// TwinCAT 3 PLC project ShowPLC
// ProgramVersion: 3.1.4026.27
// libraries:
//   Tc2_Standard, * (Beckhoff Automation GmbH)
//   Tc2_SUPS, * (Beckhoff Automation GmbH)
//   Tc2_System, * (Beckhoff Automation GmbH)
//   Tc2_Utilities, * (Beckhoff Automation GmbH)
//   Tc3_IotBase, * (Beckhoff Automation GmbH)
//   Tc3_IPCDiag, * (Beckhoff Automation GmbH)
//   Tc3_JsonXml, * (Beckhoff Automation GmbH)
// project tree:
//   DUTs/ E_JsonSection.TcDUT, E_LoadKind.TcDUT, ST_AcMeasurement.TcDUT, ST_BoxConfig.TcDUT, ST_FeedConfig.TcDUT, ST_GenericLoadConfig.TcDUT, ST_Harmonics.TcDUT, ST_LoadDemand.TcDUT, ST_MqttConfig.TcDUT
//   GVLs/ GVL_Config.TcGVL, GVL_Param.TcGVL, GVL_Persist.TcGVL
//   / PlcTask.TcTTO
//   POUs/ITFs/ I_FeedLoad.TcIO, I_JsonSource.TcIO, I_PowerMeter.TcIO
//   POUs/ MAIN.TcPOU
//   POUs/Power/ FB_EcPowerSupply.TcPOU, FB_GenericLoad.TcPOU, FB_PowerFeed.TcPOU, FB_PowerMeter_Sim.TcPOU, FB_SatelliteController.TcPOU
//   POUs/System/ FB_HostThermal.TcPOU (not stored), FB_ShowClock.TcPOU, FB_Telemetry.TcPOU, FB_IpcDiagnostics.TcPOU
//   POUs/Util/ F_CableFactor.TcPOU, F_CableLossW.TcPOU, F_CleanReal.TcPOU, F_CycleTimeS.TcPOU, F_FeedIdString.TcPOU, F_JsonHarmArray.TcPOU, F_JsonInt.TcPOU, F_JsonNum.TcPOU, F_JsonNumSigned.TcPOU, F_LowPass.TcPOU, F_PadNum.TcPOU, F_PowerAfterCable.TcPOU, F_WireOhms.TcPOU
// real-time tasks:
//   TASK PlcTask: cycle T#10ms, priority 20, ADS port 350
// I/O:
//   DEVICE Device 1 (EtherCAT), AmsNetId 192.168.30.11.2.1
//     Term 1 (EK1200) [EK1200-5000 EtherCAT Power supply (2A E-Bus)]
//       Term 10 (EL6070-0033) [EL6070-0033 1Ch. Licence key terminal, individual licences]
//       Term 2 (EL6090) [EL6090 Display terminal]
//       Term 3 (EL9227-5500) [EL9227-5500 Overcurrent protection 24V DC, 2Ch., max. 10A (sum), adjustable, extended functionalities]
//       Term 4 (EL9184) [EL9184 Potential Connection, 8 x 24V, 8 x Ground]
//       Term 5 (EL1259) [EL1259 8Ch. Dig Input 24V/8Ch. Dig. Output 24V with Multi-Time-Stamp]
//       Term 6 (EL3453-0100) [EL3453 3Ch. Power Measuring 100V]
//       Term 7 (EL3453-0100) [EL3453 3Ch. Power Measuring 100V]
//       Term 8 (EK1110) [EK1110 EtherCAT extension]
//     Box 17 (PS2001-2410) [PS2001-2410-1001 Power supply (24V, 10A, 1-phase)]
// variable links:
//   ShowPLC/ShowPLC Instance <-> Device 1 (EtherCAT)
//     PlcTask Inputs/MAIN.fbIpc.nEcCfgSlaves <-> InfoData/CfgSlaveCount
//     PlcTask Inputs/MAIN.fbIpc.nEcDevState <-> Inputs/DevState
//     PlcTask Inputs/MAIN.fbIpc.nEcSlaveCount <-> Inputs/SlaveCount

CONFIGURATION ShowPLC
    RESOURCE PLC ON TwinCAT3
        TASK PlcTask(INTERVAL := T#10ms, PRIORITY := 20);
        PROGRAM MAIN WITH PlcTask : MAIN;
    END_RESOURCE
END_CONFIGURATION

// ---- DUTs/E_JsonSection.TcDUT
{attribute 'qualified_only'}
{attribute 'strict'}
TYPE E_JsonSection :
(
    Circuit := 0,   // one row of the website's original circuits[] list
    Feed,           // one row of feeds[]
    Box,            // one row of boxes[]
    Load,           // one row of loads[]
    Diag,           // the body of the diag payload
    Harmonics       // one row of the harmonics payload
);
END_TYPE

// ---- DUTs/E_LoadKind.TcDUT
{attribute 'qualified_only'}
{attribute 'strict'}
TYPE E_LoadKind :
(
    Measured := 0,  // has its own measurement (box with an EtherCAT power supply)
    Rated,          // fixed rated power (generic load)
    Estimated       // gets a share of whatever is left on the feed (box without a supply)
);
END_TYPE

// ---- DUTs/ST_AcMeasurement.TcDUT
TYPE ST_AcMeasurement :
STRUCT
    bValid        : BOOL;   // the values below can be used
    bThdValid     : BOOL;   // the four THD values can be used
    fVoltsL1      : LREAL;  // V, L1 to ground
    fVoltsL2      : LREAL;  // V, L2 to ground
    fVoltsLL      : LREAL;  // V, L1 to L2
    fAmpsL1       : LREAL;  // A
    fAmpsL2       : LREAL;  // A
    fAmpsResidual : LREAL;  // A, summation transformer on the IN channel
    fPowerW       : LREAL;  // W,  P(L1) + P(L2)
    fApparentVA   : LREAL;  // VA, S(L1) + S(L2)
    fPowerFactor  : LREAL;  // 0..1
    fFrequencyHz  : LREAL;
    fThdVoltsL1   : LREAL;  // %
    fThdVoltsL2   : LREAL;  // %
    fThdAmpsL1    : LREAL;  // %
    fThdAmpsL2    : LREAL;  // %
END_STRUCT
END_TYPE

// ---- DUTs/ST_BoxConfig.TcDUT
TYPE ST_BoxConfig :
STRUCT
    sId               : STRING(20);     // slug of the name: lowercase letters, digits and '-'
    sControllerName   : STRING(40);     // exactly the label the website uses for this controller
    nFeedId           : INT := 1;       // index into GVL_Config.aFeeds
    bHasEcPowerSupply : BOOL;           // TRUE: live values come from the EtherCAT supply in the box
    nPixelCount       : UDINT;
    fMaxDcCurrent     : LREAL := 20.0;  // A
    fNominalDcVolts   : LREAL := 24.0;  // turns an estimated share into DC amps
    fPsuEfficiency    : LREAL := 0.95;  // DC power out / AC power in
    fWireLengthFt     : LREAL := 0.0;   // one-way length of the box's AC cable from where it branches off the feed
    nWireAwg          : INT := 12;      // AWG of one conductor, copper
END_STRUCT
END_TYPE

// ---- DUTs/ST_FeedConfig.TcDUT
TYPE ST_FeedConfig :
STRUCT
    sId           : STRING(20);     // short id used in the payloads: F1, F2
    sName         : STRING(40);
    fMaxAmps      : LREAL := 32.0;  // A per leg
    fWireLengthFt : LREAL := 0.0;   // one-way length of the infeed cable: meter to the point where the boxes branch off
    nWireAwg      : INT := 10;      // AWG of one conductor, copper
END_STRUCT
END_TYPE

// ---- DUTs/ST_GenericLoadConfig.TcDUT
TYPE ST_GenericLoadConfig :
STRUCT
    sId           : STRING(20);  // L1, L2, ...
    sName         : STRING(40);
    nFeedId       : INT := 1;    // index into GVL_Config.aFeeds
    fRatedPowerW  : LREAL;       // W at the load
    bEnabled      : BOOL;        // FALSE: counts as 0 W
    fWireLengthFt : LREAL := 0.0; // one-way length of the load's cable from where it branches off the feed
    nWireAwg      : INT := 14;   // AWG of one conductor, copper
END_STRUCT
END_TYPE

// ---- DUTs/ST_Harmonics.TcDUT
TYPE ST_Harmonics :
STRUCT
    bValid   : BOOL;
    aVoltsL1 : ARRAY[2..GVL_Param.HARMONIC_MAX_ORDER] OF LREAL;
    aVoltsL2 : ARRAY[2..GVL_Param.HARMONIC_MAX_ORDER] OF LREAL;
    aAmpsL1  : ARRAY[2..GVL_Param.HARMONIC_MAX_ORDER] OF LREAL;
    aAmpsL2  : ARRAY[2..GVL_Param.HARMONIC_MAX_ORDER] OF LREAL;
END_STRUCT
END_TYPE

// ---- DUTs/ST_LoadDemand.TcDUT
TYPE ST_LoadDemand :
STRUCT
    eKind        : E_LoadKind;  // how the feed treats this load
    fAcPowerW    : LREAL;       // W the load takes at the branch point, its own cable loss included. Measured and Rated loads only
    fCableLossW  : LREAL;       // W lost in the load's own cable. Measured and Rated: part of fAcPowerW. Estimated: from its current share
    fWeight      : LREAL;       // share weight: the pixel count. Estimated loads only
    fCableFactor : LREAL;       // 1/W: loss in the load's own cable = fCableFactor * (power at the load)^2. Estimated loads only
    bValid       : BOOL;        // FALSE: a measured load that is not reporting
END_STRUCT
END_TYPE

// ---- DUTs/ST_MqttConfig.TcDUT
TYPE ST_MqttConfig :
STRUCT
    bEnable     : BOOL := TRUE;
    sHost       : STRING(63) := '192.168.30.31';
    nPort       : UINT := 1883;
    sClientId   : STRING(63) := 'sfl-plc';
    sUser       : STRING(63) := 'plc';
    nKeepAliveS : UINT := 30;
    sTopicRoot  : STRING(63) := 'sfl/plc';
    tDashboard  : TIME := T#1S;
    tDiag       : TIME := T#5S;
    tHarmonics  : TIME := T#10S;
END_STRUCT
END_TYPE

// ---- GVLs/GVL_Config.TcGVL
{attribute 'qualified_only'}
VAR_GLOBAL
    // ---- development switches -------------------------------------------------
    bSimulateMeters   : BOOL := TRUE;   // TRUE: feeds read FB_PowerMeter_Sim. Set FALSE in step 4
    bSimulateSupplies : BOOL := TRUE;   // TRUE: supplies use their fSim values. Set FALSE in step 5

    // ---- model ----------------------------------------------------------------
    fFilterTimeS      : LREAL := 1.0;   // low-pass on feed and supply values before the split, seconds
    fVoltsPresentMin  : LREAL := 90.0;  // V per leg. Above this a feed counts as "on"

    // ---- cables ---------------------------------------------------------------
    // Every feed, box and load has a one-way cable length and an AWG. The loss in each cable is I^2 R
    // with that component's own current. Lengths below are placeholders until measured.
    fWireTempC          : LREAL := 20.0;   // conductor temperature for the resistance. Copper: +0.39 % per degree C
    fWireFactor         : LREAL := 1.0;    // 1.0 solid copper, about 1.03 stranded copper, about 1.6 aluminium
    fNominalAcVolts     : LREAL := 240.0;  // L1 to L2 at the loads. With the power factor it turns a load's power into the current in its cable
    fNominalPowerFactor : LREAL := 1.0;    // of the boxes and loads. Current = power / (volts * power factor)

    // ---- feeds ----------------------------------------------------------------
    aFeeds : ARRAY[1..GVL_Param.FEED_COUNT] OF ST_FeedConfig := [
        (sId := 'F1', sName := 'Feed 1', fMaxAmps := 32.0, fWireLengthFt := 100.0, nWireAwg := 10),
        (sId := 'F2', sName := 'Feed 2', fMaxAmps := 32.0, fWireLengthFt := 100.0, nWireAwg := 10)];

    // ---- satellite controller boxes ---------------------------------------------
    // sControllerName must match the website's label exactly. sId is its slug.
    // A box without an EtherCAT supply is estimated from its feed. Its DC amps use fNominalDcVolts (24 V unless set here).
    aBoxes : ARRAY[1..GVL_Param.BOX_COUNT] OF ST_BoxConfig := [
        (sId := 'porch',        sControllerName := 'Porch',        nFeedId := 1, bHasEcPowerSupply := FALSE, nPixelCount := 16325, fMaxDcCurrent := 80.0, fWireLengthFt := 50.0, nWireAwg := 12),
        (sId := 'metal-roof',   sControllerName := 'Metal Roof',   nFeedId := 2, bHasEcPowerSupply := FALSE, nPixelCount := 12820, fMaxDcCurrent := 80.0, fWireLengthFt := 50.0, nWireAwg := 12),
        (sId := 'center-gable', sControllerName := 'Center Gable', nFeedId := 1, bHasEcPowerSupply := TRUE,  nPixelCount := 2841,  fMaxDcCurrent := 20.0, fWireLengthFt := 50.0, nWireAwg := 12),
        (sId := 'courtyard',    sControllerName := 'Courtyard',    nFeedId := 1, bHasEcPowerSupply := TRUE,  nPixelCount := 452,   fMaxDcCurrent := 20.0, fWireLengthFt := 50.0, nWireAwg := 12),
        (sId := 'lawn-s-1',     sControllerName := 'Lawn S-1',     nFeedId := 1, bHasEcPowerSupply := TRUE,  nPixelCount := 1500,  fMaxDcCurrent := 20.0, fWireLengthFt := 50.0, nWireAwg := 12),
        (sId := 'lawn-s-2',     sControllerName := 'Lawn S-2',     nFeedId := 1, bHasEcPowerSupply := TRUE,  nPixelCount := 2541,  fMaxDcCurrent := 20.0, fWireLengthFt := 50.0, nWireAwg := 12),
        (sId := 'lawn-s-3',     sControllerName := 'Lawn S-3',     nFeedId := 2, bHasEcPowerSupply := TRUE,  nPixelCount := 6141,  fMaxDcCurrent := 20.0, fWireLengthFt := 50.0, nWireAwg := 12),
        (sId := 'lawn-n-1',     sControllerName := 'Lawn N-1',     nFeedId := 2, bHasEcPowerSupply := TRUE,  nPixelCount := 2450,  fMaxDcCurrent := 20.0, fWireLengthFt := 50.0, nWireAwg := 12),
        (sId := 'lawn-n-2',     sControllerName := 'Lawn N-2',     nFeedId := 2, bHasEcPowerSupply := TRUE,  nPixelCount := 4115,  fMaxDcCurrent := 20.0, fWireLengthFt := 50.0, nWireAwg := 12)];

    // ---- generic loads ------------------------------------------------------------
    // One row per GVL_Param.LOAD_COUNT.
    aLoads : ARRAY[1..GVL_Param.LOAD_COUNT] OF ST_GenericLoadConfig := [
        (sId := 'L1', sName := 'Metal Roof Floods', nFeedId := 2, fRatedPowerW := 20.0, bEnabled := TRUE, fWireLengthFt := 50.0, nWireAwg := 14),
        (sId := 'L2', sName := 'North Peak Floods', nFeedId := 2, fRatedPowerW := 20.0, bEnabled := TRUE, fWireLengthFt := 50.0, nWireAwg := 14),
        (sId := 'L3', sName := 'South Peak Floods', nFeedId := 2, fRatedPowerW := 20.0, bEnabled := TRUE, fWireLengthFt := 50.0, nWireAwg := 14)];

    // ---- EtherCAT power supplies (PS2001) -------------------------------------------
    // Info data scaling is not documented. 0.0 keeps the value out of the payload until it is checked in step 5.
    fPsuInfo1Scale : LREAL := 0.0;      // degrees C per count of "Info data 1" (temperature)
    fPsuInfo2Scale : LREAL := 0.0;      // volts per count of "Info data 2" (RMS input voltage)

    // ---- TF8330 -----------------------------------------------------------------------
    nTf8330FundamentalIndex : INT := 1; // element of aHarm1 that reads 100 (the fundamental): 1 if element 0 is the DC part, 0 if the arrays start at the fundamental, -1 if they start at the 2nd harmonic. Check in step 4

    // ---- MQTT ---------------------------------------------------------------------------
    stMqtt : ST_MqttConfig;             // defaults are in the type

    // ---- local time, for the midnight energy reset: US Central ---------------------------
    // UTC = local time + bias (minutes). wDay is the occurrence in the month: 1 = first, 2 = second, 5 = last.
    stTimeZone : ST_TimeZoneInformation := (
        bias         := 360,
        standardName := 'CST',
        standardDate := (wYear := 0, wMonth := 11, wDayOfWeek := 0, wDay := 1, wHour := 2),
        standardBias := 0,
        daylightName := 'CDT',
        daylightDate := (wYear := 0, wMonth := 3, wDayOfWeek := 0, wDay := 2, wHour := 2),
        daylightBias := -60);
END_VAR

// ---- GVLs/GVL_Param.TcGVL
{attribute 'qualified_only'}
VAR_GLOBAL CONSTANT
    FEED_COUNT         : INT := 2;
    BOX_COUNT          : INT := 9;
    LOAD_COUNT         : INT := 3;
    MAX_LOADS_PER_FEED : INT := GVL_Param.BOX_COUNT + GVL_Param.LOAD_COUNT;
    HARMONIC_MAX_ORDER : INT := 25;  // highest harmonic order kept and published. 2..63
END_VAR

// ---- GVLs/GVL_Persist.TcGVL
{attribute 'qualified_only'}
VAR_GLOBAL PERSISTENT
    sMqttPassword : STRING(63);                                  // empty = telemetry stays offline
    aEnergyWh     : ARRAY[1..GVL_Param.FEED_COUNT] OF LREAL;     // Wh per feed since local midnight
    nEnergyDay    : UDINT;                                       // local day number the counters belong to
END_VAR

// ---- POUs/ITFs/I_FeedLoad.TcIO
INTERFACE I_FeedLoad

// What this load asks of its feed this cycle.
METHOD GetDemand : ST_LoadDemand
END_METHOD

// The feed's answer to an Estimated load: its share of the unmeasured power.
METHOD SetShare
VAR_INPUT
    fShareW     : LREAL;  // W on the AC side
    bShareValid : BOOL;   // FALSE: the feed has no valid measurement
END_VAR
END_METHOD

END_INTERFACE

// ---- POUs/ITFs/I_JsonSource.TcIO
INTERFACE I_JsonSource

// Writes the keys of one JSON object. The caller opens and closes the object.
METHOD WriteJson
VAR_INPUT
    eSection : E_JsonSection;
END_VAR
VAR_IN_OUT
    fbJson : FB_JsonSaxWriter;
END_VAR
END_METHOD

END_INTERFACE

// ---- POUs/ITFs/I_PowerMeter.TcIO
INTERFACE I_PowerMeter

// Fills stMeas. Returns TRUE when the values are valid.
METHOD Read : BOOL
VAR_IN_OUT
    stMeas : ST_AcMeasurement;
END_VAR
END_METHOD

// Fills stHarm. Returns TRUE when the values are valid.
METHOD ReadHarmonics : BOOL
VAR_IN_OUT
    stHarm : ST_Harmonics;
END_VAR
END_METHOD

END_INTERFACE

// ---- POUs/MAIN.TcPOU
PROGRAM MAIN
VAR
    // Power model
    aFeeds     : ARRAY[1..GVL_Param.FEED_COUNT] OF FB_PowerFeed;
    aSimMeters : ARRAY[1..GVL_Param.FEED_COUNT] OF FB_PowerMeter_Sim;
    aBoxes     : ARRAY[1..GVL_Param.BOX_COUNT] OF FB_SatelliteController;
    aLoads     : ARRAY[1..GVL_Param.LOAD_COUNT] OF FB_GenericLoad;
    ipMeter    : I_PowerMeter;

    // Totals for the website's top-level keys
    fTotalPowerW   : LREAL;
    fTotalAmps     : LREAL;
    fEnergyTodayWh : LREAL;

    // Reporting
    fbClock     : FB_ShowClock;
    fbTelemetry : FB_Telemetry;
    fbIpc       : FB_IpcDiagnostics;

    // Persistent data
    bSavePersistent : BOOL;                    // set TRUE online to store GVL_Persist now
    fbSavePersist   : FB_WritePersistentData;

    i : INT;
    n : INT;
END_VAR

// Clock. On a new local day the energy counters start again
fbClock();
IF fbClock.bValid AND (fbClock.nLocalDay <> GVL_Persist.nEnergyDay) THEN
    FOR i := 1 TO GVL_Param.FEED_COUNT DO
        GVL_Persist.aEnergyWh[i] := 0.0;
    END_FOR
    GVL_Persist.nEnergyDay := fbClock.nLocalDay;
END_IF

// Feeds: read the meter, filter, cable loss, start a new load list
FOR i := 1 TO GVL_Param.FEED_COUNT DO
    ipMeter := aSimMeters[i];
    aFeeds[i](stCfg := GVL_Config.aFeeds[i], ipMeter := ipMeter, fEnergyWh := GVL_Persist.aEnergyWh[i]);
END_FOR

// Boxes and generic loads: update, then report to their feed
FOR i := 1 TO GVL_Param.BOX_COUNT DO
    aBoxes[i](stCfg := GVL_Config.aBoxes[i]);
    n := GVL_Config.aBoxes[i].nFeedId;
    IF (n >= 1) AND (n <= GVL_Param.FEED_COUNT) THEN
        aFeeds[n].AddLoad(ipLoad := aBoxes[i]);
    ELSE
        aBoxes[i].SetShare(fShareW := 0.0, bShareValid := FALSE);  // nFeedId names no feed: nothing to estimate from
    END_IF
END_FOR
FOR i := 1 TO GVL_Param.LOAD_COUNT DO
    aLoads[i](stCfg := GVL_Config.aLoads[i]);
    n := GVL_Config.aLoads[i].nFeedId;
    IF (n >= 1) AND (n <= GVL_Param.FEED_COUNT) THEN
        aFeeds[n].AddLoad(ipLoad := aLoads[i]);
    END_IF
END_FOR

// Feeds: split what is left between the boxes without a supply, and add up the totals
fTotalPowerW   := 0.0;
fTotalAmps     := 0.0;
fEnergyTodayWh := 0.0;
FOR i := 1 TO GVL_Param.FEED_COUNT DO
    aFeeds[i].Allocate();
    IF aFeeds[i].bValid THEN
        fTotalPowerW := fTotalPowerW + MAX(0.0, aFeeds[i].stMeas.fPowerW);
        fTotalAmps   := fTotalAmps + aFeeds[i].fAmps;
    END_IF
    fEnergyTodayWh := fEnergyTodayWh + GVL_Persist.aEnergyWh[i];
END_FOR

// Controller health
fbIpc();

// Telemetry: hand over the sources, then let it publish
FOR i := 1 TO GVL_Param.FEED_COUNT DO
    fbTelemetry.AddSource(eSection := E_JsonSection.Feed, ipSource := aFeeds[i]);
END_FOR
FOR i := 1 TO GVL_Param.BOX_COUNT DO
    fbTelemetry.AddSource(eSection := E_JsonSection.Box, ipSource := aBoxes[i]);
END_FOR
FOR i := 1 TO GVL_Param.LOAD_COUNT DO
    fbTelemetry.AddSource(eSection := E_JsonSection.Load, ipSource := aLoads[i]);
END_FOR
fbTelemetry.AddSource(eSection := E_JsonSection.Diag, ipSource := fbIpc);
fbTelemetry(stCfg := GVL_Config.stMqtt, sPassword := GVL_Persist.sMqttPassword, sTimestamp := fbClock.sUtcIso,
            bSimulated := GVL_Config.bSimulateMeters OR GVL_Config.bSimulateSupplies,
            fTotalPowerW := fTotalPowerW, fTotalAmps := fTotalAmps, fEnergyTodayWh := fEnergyTodayWh);

// Store GVL_Persist on request: set bSavePersistent to TRUE online, once
fbSavePersist(NETID := '', PORT := _AppInfo.AdsPort, START := bSavePersistent, TMOUT := T#5S);
bSavePersistent := FALSE;

END_PROGRAM

// ---- POUs/Power/FB_PowerFeed.TcPOU
FUNCTION_BLOCK FB_PowerFeed IMPLEMENTS I_JsonSource
VAR_INPUT
    stCfg   : ST_FeedConfig;  // this feed's row of GVL_Config.aFeeds
    ipMeter : I_PowerMeter;   // where the measurement comes from
END_VAR
VAR_IN_OUT
    fEnergyWh : LREAL;        // energy counter owned by the caller (persistent)
END_VAR
VAR_OUTPUT
    bValid         : BOOL;              // the meter delivers valid data
    bDegraded      : BOOL;              // a box with a supply on this feed is not reporting: estimates are too high
    stMeas         : ST_AcMeasurement;  // filtered measurement
    fAmps          : LREAL;             // A, the larger leg
    fCableLossW    : LREAL;             // W lost in the infeed cable
    fLoadPowerW    : LREAL;             // W at the branch point: meter minus infeed cable loss
    fMeasuredW     : LREAL;             // W taken by boxes with a supply, their cable losses included
    fRatedW        : LREAL;             // W taken by enabled generic loads, their cable losses included
    fUnmeteredW    : LREAL;             // W split across boxes without a supply, their cable losses included
    fDropLossW     : LREAL;             // W lost in the loads' own cables, as the loads report it
    fUnaccountedW  : LREAL;             // W left over. Not zero means the model is off
    fEnergyTodayWh : LREAL;             // copy of the counter for telemetry
    nLoadCount     : INT;               // loads registered this cycle
END_VAR
VAR
    stRaw     : ST_AcMeasurement;
    aLoads    : ARRAY[1..GVL_Param.MAX_LOADS_PER_FEED] OF I_FeedLoad;
    bMeterOk  : BOOL;
    fCycleS   : LREAL;
    fTau      : LREAL;
    fOhms     : LREAL;
    fRawLossW : LREAL;  // infeed loss from this cycle's unfiltered currents
END_VAR

fCycleS := F_CycleTimeS();
fTau    := GVL_Config.fFilterTimeS;

// 1. Read the meter
bMeterOk := FALSE;
IF ipMeter <> 0 THEN
    bMeterOk := ipMeter.Read(stMeas := stRaw);
END_IF

// 2. Infeed cable loss from the raw leg currents. The ground conductor carries no load current, so two conductors count.
//    The loss goes with the square of the current, so it is computed before the filter and filtered on its own:
//    squaring a filtered current would read low whenever the load moves.
fOhms     := F_WireOhms(fLengthFt := stCfg.fWireLengthFt, nAwg := stCfg.nWireAwg);
fRawLossW := fOhms * (stRaw.fAmpsL1 * stRaw.fAmpsL1 + stRaw.fAmpsL2 * stRaw.fAmpsL2);

// 3. Filter what the power balance uses. Everything else is passed through.
IF bMeterOk THEN
    IF bValid THEN
        stRaw.fAmpsL1       := F_LowPass(fState := stMeas.fAmpsL1,       fInput := stRaw.fAmpsL1,       fTimeS := fTau, fCycleS := fCycleS);
        stRaw.fAmpsL2       := F_LowPass(fState := stMeas.fAmpsL2,       fInput := stRaw.fAmpsL2,       fTimeS := fTau, fCycleS := fCycleS);
        stRaw.fAmpsResidual := F_LowPass(fState := stMeas.fAmpsResidual, fInput := stRaw.fAmpsResidual, fTimeS := fTau, fCycleS := fCycleS);
        stRaw.fPowerW       := F_LowPass(fState := stMeas.fPowerW,       fInput := stRaw.fPowerW,       fTimeS := fTau, fCycleS := fCycleS);
        stRaw.fApparentVA   := F_LowPass(fState := stMeas.fApparentVA,   fInput := stRaw.fApparentVA,   fTimeS := fTau, fCycleS := fCycleS);
        fCableLossW         := F_LowPass(fState := fCableLossW,          fInput := fRawLossW,           fTimeS := fTau, fCycleS := fCycleS);
    ELSE
        fCableLossW := fRawLossW;
    END_IF
    stMeas := stRaw;  // on the first valid sample this is the raw value: no filter run-in
END_IF
bValid := bMeterOk;
stMeas.bValid := bMeterOk;

fAmps := MAX(stMeas.fAmpsL1, stMeas.fAmpsL2);
fLoadPowerW := MAX(0.0, stMeas.fPowerW - fCableLossW);

// 4. Energy since local midnight. TF8330 has no energy counters, so it is integrated here.
IF bValid THEN
    fEnergyWh := fEnergyWh + MAX(0.0, stMeas.fPowerW) * fCycleS / 3600.0;
END_IF
fEnergyTodayWh := fEnergyWh;

// 5. New load list. MAIN hands every load in again each cycle, so no reference outlives a cycle.
nLoadCount := 0;

// Registers a load for this cycle. Returns FALSE when the list is full.
METHOD AddLoad : BOOL
VAR_INPUT
    ipLoad : I_FeedLoad;
END_VAR
AddLoad := FALSE;
IF (ipLoad <> 0) AND (nLoadCount < GVL_Param.MAX_LOADS_PER_FEED) THEN
    nLoadCount := nLoadCount + 1;
    aLoads[nLoadCount] := ipLoad;
    AddLoad := TRUE;
END_IF
END_METHOD

// Call once per cycle after every load has been added.
METHOD Allocate
VAR
    i          : INT;
    stDemand   : ST_LoadDemand;
    fWeightSum : LREAL;  // sum of the pixel counts of the estimated boxes
    fFactorSum : LREAL;  // sum of (cable factor * pixel count^2) over them
    fRest      : LREAL;  // W left for them, at the branch point
    fPerPixel  : LREAL;  // W per pixel at the boxes
    fAtBox     : LREAL;
    fShare     : LREAL;
END_VAR
fMeasuredW := 0.0;
fRatedW    := 0.0;
fDropLossW := 0.0;
fWeightSum := 0.0;
fFactorSum := 0.0;
bDegraded  := FALSE;

// Pass 1: add up what is known. Every demand is at the branch point, cable loss included.
FOR i := 1 TO nLoadCount DO
    stDemand := aLoads[i].GetDemand();
    CASE stDemand.eKind OF
        E_LoadKind.Measured:
            IF stDemand.bValid THEN
                fMeasuredW := fMeasuredW + MAX(0.0, stDemand.fAcPowerW);
                fDropLossW := fDropLossW + MAX(0.0, stDemand.fCableLossW);
            ELSE
                bDegraded := TRUE;
            END_IF
        E_LoadKind.Rated:
            fRatedW    := fRatedW + MAX(0.0, stDemand.fAcPowerW);
            fDropLossW := fDropLossW + MAX(0.0, stDemand.fCableLossW);
        E_LoadKind.Estimated:
            fWeightSum := fWeightSum + MAX(0.0, stDemand.fWeight);
            fFactorSum := fFactorSum + MAX(0.0, stDemand.fCableFactor) * stDemand.fWeight * stDemand.fWeight;
    END_CASE
END_FOR

// What is left for the boxes without a supply
fRest := MAX(0.0, fLoadPowerW - fMeasuredW - fRatedW);
IF fWeightSum > 0.0 THEN
    fUnmeteredW := fRest;
ELSE
    fUnmeteredW := 0.0;
END_IF
fUnaccountedW := fLoadPowerW - fMeasuredW - fRatedW - fUnmeteredW;

// The split is proportional to pixels AT THE BOXES: box i gets fPerPixel * pixels at its terminals and takes
// that plus its own cable loss, a_i * (fPerPixel * pixels)^2, at the branch point. The sum over the boxes
// equals fRest, which gives fPerPixel from a quadratic: fFactorSum * k^2 + fWeightSum * k = fRest.
fPerPixel := 0.0;
IF fWeightSum > 0.0 THEN
    fPerPixel := 2.0 * fRest / (fWeightSum + SQRT(fWeightSum * fWeightSum + 4.0 * fFactorSum * fRest));
END_IF

// Pass 2: hand out the shares at the branch point; each box recovers its own power from its share.
FOR i := 1 TO nLoadCount DO
    stDemand := aLoads[i].GetDemand();
    IF stDemand.eKind = E_LoadKind.Estimated THEN
        fAtBox := fPerPixel * MAX(0.0, stDemand.fWeight);
        fShare := fAtBox + MAX(0.0, stDemand.fCableFactor) * fAtBox * fAtBox;
        aLoads[i].SetShare(fShareW := fShare, bShareValid := bValid);
        stDemand   := aLoads[i].GetDemand();  // now carries this cycle's cable loss
        fDropLossW := fDropLossW + MAX(0.0, stDemand.fCableLossW);
    END_IF
END_FOR
END_METHOD

METHOD WriteJson
VAR_INPUT
    eSection : E_JsonSection;
END_VAR
VAR_IN_OUT
    fbJson : FB_JsonSaxWriter;
END_VAR
VAR
    bLegsLive : BOOL;
    bThdOk    : BOOL;
    bHarmOk   : BOOL;
    stHarm    : ST_Harmonics;
END_VAR
CASE eSection OF

    E_JsonSection.Circuit:
        bLegsLive := bValid AND (stMeas.fVoltsL1 > GVL_Config.fVoltsPresentMin) AND (stMeas.fVoltsL2 > GVL_Config.fVoltsPresentMin);
        fbJson.AddKey('id');
        fbJson.AddString(stCfg.sId);
        fbJson.AddKey('name');
        fbJson.AddString(stCfg.sName);
        fbJson.AddKey('on');
        fbJson.AddBool(bLegsLive);
        F_JsonNum(sKey := 'amps', fValue := fAmps, bValid := bValid, nDecimals := 2, fbJson := fbJson);

    E_JsonSection.Feed:
        bThdOk := bValid AND stMeas.bThdValid;
        fbJson.AddKey('id');
        fbJson.AddString(stCfg.sId);
        fbJson.AddKey('name');
        fbJson.AddString(stCfg.sName);
        fbJson.AddKey('ok');
        fbJson.AddBool(bValid);
        fbJson.AddKey('degraded');
        fbJson.AddBool(bDegraded);
        F_JsonNum(sKey := 'maxAmps',       fValue := stCfg.fMaxAmps,         bValid := TRUE,   nDecimals := 1, fbJson := fbJson);
        F_JsonNum(sKey := 'amps',          fValue := fAmps,                  bValid := bValid, nDecimals := 2, fbJson := fbJson);
        F_JsonNum(sKey := 'ampsL1',        fValue := stMeas.fAmpsL1,         bValid := bValid, nDecimals := 2, fbJson := fbJson);
        F_JsonNum(sKey := 'ampsL2',        fValue := stMeas.fAmpsL2,         bValid := bValid, nDecimals := 2, fbJson := fbJson);
        F_JsonNum(sKey := 'ampsResidual',  fValue := stMeas.fAmpsResidual,   bValid := bValid, nDecimals := 3, fbJson := fbJson);
        F_JsonNum(sKey := 'voltsL1',       fValue := stMeas.fVoltsL1,        bValid := bValid, nDecimals := 1, fbJson := fbJson);
        F_JsonNum(sKey := 'voltsL2',       fValue := stMeas.fVoltsL2,        bValid := bValid, nDecimals := 1, fbJson := fbJson);
        F_JsonNum(sKey := 'voltsLL',       fValue := stMeas.fVoltsLL,        bValid := bValid, nDecimals := 1, fbJson := fbJson);
        F_JsonNum(sKey := 'powerW',        fValue := stMeas.fPowerW,         bValid := bValid, nDecimals := 1, fbJson := fbJson);
        F_JsonNum(sKey := 'apparentVA',    fValue := stMeas.fApparentVA,     bValid := bValid, nDecimals := 1, fbJson := fbJson);
        F_JsonNum(sKey := 'pf',            fValue := stMeas.fPowerFactor,    bValid := bValid, nDecimals := 2, fbJson := fbJson);
        F_JsonNum(sKey := 'hz',            fValue := stMeas.fFrequencyHz,    bValid := bValid, nDecimals := 2, fbJson := fbJson);
        F_JsonNum(sKey := 'thdVoltsL1',    fValue := stMeas.fThdVoltsL1,     bValid := bThdOk, nDecimals := 1, fbJson := fbJson);
        F_JsonNum(sKey := 'thdVoltsL2',    fValue := stMeas.fThdVoltsL2,     bValid := bThdOk, nDecimals := 1, fbJson := fbJson);
        F_JsonNum(sKey := 'thdAmpsL1',     fValue := stMeas.fThdAmpsL1,      bValid := bThdOk, nDecimals := 1, fbJson := fbJson);
        F_JsonNum(sKey := 'thdAmpsL2',     fValue := stMeas.fThdAmpsL2,      bValid := bThdOk, nDecimals := 1, fbJson := fbJson);
        F_JsonNum(sKey := 'cableLossW',    fValue := fCableLossW,            bValid := bValid, nDecimals := 1, fbJson := fbJson);
        F_JsonNum(sKey := 'dropLossW',     fValue := fDropLossW,             bValid := bValid, nDecimals := 1, fbJson := fbJson);
        F_JsonNum(sKey := 'measuredW',     fValue := fMeasuredW,             bValid := bValid, nDecimals := 1, fbJson := fbJson);
        F_JsonNum(sKey := 'ratedW',        fValue := fRatedW,                bValid := TRUE,   nDecimals := 1, fbJson := fbJson);
        F_JsonNum(sKey := 'unmeteredW',    fValue := fUnmeteredW,            bValid := bValid, nDecimals := 1, fbJson := fbJson);
        F_JsonNumSigned(sKey := 'unaccountedW', fValue := fUnaccountedW,     bValid := bValid, nDecimals := 1, fbJson := fbJson);
        F_JsonNum(sKey := 'energyTodayWh', fValue := fEnergyTodayWh,         bValid := TRUE,   nDecimals := 0, fbJson := fbJson);

    E_JsonSection.Harmonics:
        bHarmOk := FALSE;
        IF ipMeter <> 0 THEN
            bHarmOk := ipMeter.ReadHarmonics(stHarm := stHarm);
        END_IF
        fbJson.AddKey('id');
        fbJson.AddString(stCfg.sId);
        fbJson.AddKey('ok');
        fbJson.AddBool(bHarmOk);
        F_JsonHarmArray(sKey := 'ampsL1',  bValid := bHarmOk, fbJson := fbJson, aValues := stHarm.aAmpsL1);
        F_JsonHarmArray(sKey := 'ampsL2',  bValid := bHarmOk, fbJson := fbJson, aValues := stHarm.aAmpsL2);
        F_JsonHarmArray(sKey := 'voltsL1', bValid := bHarmOk, fbJson := fbJson, aValues := stHarm.aVoltsL1);
        F_JsonHarmArray(sKey := 'voltsL2', bValid := bHarmOk, fbJson := fbJson, aValues := stHarm.aVoltsL2);

END_CASE
END_METHOD

END_FUNCTION_BLOCK

// ---- POUs/Util/F_CycleTimeS.TcPOU
FUNCTION F_CycleTimeS : LREAL
VAR
    nIdx : DINT;
END_VAR

F_CycleTimeS := 0.010;  // fallback: 10 ms
nIdx := GETCURTASKINDEXEX();
IF (nIdx >= 1) AND (nIdx <= 20) THEN
    IF _TaskInfo[nIdx].CycleTime > 0 THEN
        F_CycleTimeS := UDINT_TO_LREAL(_TaskInfo[nIdx].CycleTime) * 1.0E-7;  // CycleTime is in 100 ns
    END_IF
END_IF

END_FUNCTION

// ---- POUs/Util/F_WireOhms.TcPOU
FUNCTION F_WireOhms : LREAL
VAR_INPUT
    fLengthFt : LREAL;  // one-way length of the run
    nAwg      : INT;    // AWG of one conductor. 0 = 1/0, -1 = 2/0, -2 = 3/0, -3 = 4/0
END_VAR
VAR
    fAwg       : LREAL;
    fCmil      : LREAL;  // cross-section in circular mils
    fOhmPerKft : LREAL;
    fTempC     : LREAL;
END_VAR

fAwg       := INT_TO_LREAL(LIMIT(-3, nAwg, 30));                          // 4/0 to 30 AWG. Anything else is a typo
fTempC     := LIMIT(-60.0, GVL_Config.fWireTempC, 150.0);
fCmil      := 25.0 * EXPT(92.0, (36.0 - fAwg) * 2.0 / 39.0);
fOhmPerKft := 10371.0 / fCmil * (1.0 + 0.00393 * (fTempC - 20.0)) * MAX(0.1, GVL_Config.fWireFactor);
F_WireOhms := MAX(0.0, fLengthFt) * fOhmPerKft / 1000.0;

END_FUNCTION

// ---- POUs/Util/F_LowPass.TcPOU
FUNCTION F_LowPass : LREAL
VAR_INPUT
    fState  : LREAL;  // filtered value from the previous cycle
    fInput  : LREAL;  // new raw value
    fTimeS  : LREAL;  // time constant in seconds. 0 switches the filter off
    fCycleS : LREAL;  // task cycle time in seconds
END_VAR
VAR
    fAlpha : LREAL;
END_VAR

IF (fTimeS <= 0.0) OR (fCycleS <= 0.0) THEN
    F_LowPass := fInput;
ELSE
    fAlpha := fCycleS / (fTimeS + fCycleS);
    F_LowPass := fState + fAlpha * (fInput - fState);
END_IF

END_FUNCTION

// ---- POUs/Util/F_JsonNum.TcPOU
FUNCTION F_JsonNum : BOOL
VAR_INPUT
    sKey      : STRING(31);
    fValue    : LREAL;
    bValid    : BOOL;
    nDecimals : INT;  // 0..3
END_VAR
VAR_IN_OUT
    fbJson : FB_JsonSaxWriter;
END_VAR
VAR
    fTmp   : LREAL;
    fScale : LREAL;
    bOk    : BOOL;
END_VAR

fTmp := fValue;
bOk := FALSE;
IF bValid THEN
    IF IsFinite(F_LREAL(fTmp)) THEN
        bOk := ABS(fTmp) < 1.0E12;
    END_IF
END_IF

fbJson.AddKey(sKey);
IF bOk THEN
    CASE nDecimals OF
        1: fScale := 10.0;
        2: fScale := 100.0;
        3: fScale := 1000.0;
    ELSE
        fScale := 1.0;
    END_CASE
    fTmp := LINT_TO_LREAL(LREAL_TO_LINT(fTmp * fScale)) / fScale;
    IF fTmp < 0.0 THEN
        fTmp := 0.0;
    END_IF
    fbJson.AddLreal(fTmp);
ELSE
    fbJson.AddNull();
END_IF
F_JsonNum := bOk;

END_FUNCTION

// ---- POUs/Util/F_JsonNumSigned.TcPOU
FUNCTION F_JsonNumSigned : BOOL
VAR_INPUT
    sKey      : STRING(31);
    fValue    : LREAL;
    bValid    : BOOL;
    nDecimals : INT;  // 0..3
END_VAR
VAR_IN_OUT
    fbJson : FB_JsonSaxWriter;
END_VAR
VAR
    fTmp   : LREAL;
    fScale : LREAL;
    bOk    : BOOL;
END_VAR

fTmp := fValue;
bOk := FALSE;
IF bValid THEN
    IF IsFinite(F_LREAL(fTmp)) THEN
        bOk := ABS(fTmp) < 1.0E12;
    END_IF
END_IF

fbJson.AddKey(sKey);
IF bOk THEN
    CASE nDecimals OF
        1: fScale := 10.0;
        2: fScale := 100.0;
        3: fScale := 1000.0;
    ELSE
        fScale := 1.0;
    END_CASE
    fbJson.AddLreal(LINT_TO_LREAL(LREAL_TO_LINT(fTmp * fScale)) / fScale);
ELSE
    fbJson.AddNull();
END_IF
F_JsonNumSigned := bOk;

END_FUNCTION

// ---- POUs/Util/F_JsonHarmArray.TcPOU
FUNCTION F_JsonHarmArray : BOOL
VAR_INPUT
    sKey   : STRING(31);
    bValid : BOOL;
END_VAR
VAR_IN_OUT
    fbJson  : FB_JsonSaxWriter;
    aValues : ARRAY[2..GVL_Param.HARMONIC_MAX_ORDER] OF LREAL;
END_VAR
VAR
    n  : INT;
    fV : LREAL;
END_VAR

fbJson.AddKey(sKey);
fbJson.StartArray();
IF bValid THEN
    FOR n := 2 TO GVL_Param.HARMONIC_MAX_ORDER DO
        fV := aValues[n];
        IF IsFinite(F_LREAL(fV)) THEN
            fV := LIMIT(0.0, fV, 1000.0);
            fbJson.AddLreal(LINT_TO_LREAL(LREAL_TO_LINT(fV * 10.0)) / 10.0);
        ELSE
            fbJson.AddNull();
        END_IF
    END_FOR
END_IF
fbJson.EndArray();
F_JsonHarmArray := bValid;

END_FUNCTION

// ---- POUs/Power/FB_PowerMeter_Sim.TcPOU
FUNCTION_BLOCK FB_PowerMeter_Sim IMPLEMENTS I_PowerMeter
VAR_INPUT
    bOnline      : BOOL := TRUE;    // FALSE simulates a dead meter
    fVoltsLeg    : LREAL := 120.0;  // V, each leg to ground
    fPowerW      : LREAL := 1500.0; // W, total active power of the feed
    fPowerFactor : LREAL := 0.98;
    fResidualA   : LREAL := 0.0;    // A
    fThdVoltsPct : LREAL := 2.0;
    fThdAmpsPct  : LREAL := 11.0;
END_VAR

// Nothing to do here. The feed calls Read() and ReadHarmonics().
;

METHOD Read : BOOL
VAR_IN_OUT
    stMeas : ST_AcMeasurement;
END_VAR
VAR
    fPf : LREAL;
    fVa : LREAL;
END_VAR
fPf := LIMIT(0.1, fPowerFactor, 1.0);
fVa := MAX(0.0, fPowerW) / fPf;

stMeas.bValid        := bOnline;
stMeas.bThdValid     := bOnline;
stMeas.fVoltsL1      := fVoltsLeg;
stMeas.fVoltsL2      := fVoltsLeg;
stMeas.fVoltsLL      := 2.0 * fVoltsLeg;
IF fVoltsLeg > 1.0 THEN
    stMeas.fAmpsL1 := fVa / (2.0 * fVoltsLeg);
ELSE
    stMeas.fAmpsL1 := 0.0;
END_IF
stMeas.fAmpsL2       := stMeas.fAmpsL1;
stMeas.fAmpsResidual := MAX(0.0, fResidualA);
stMeas.fPowerW       := MAX(0.0, fPowerW);
stMeas.fApparentVA   := fVa;
stMeas.fPowerFactor  := fPf;
stMeas.fFrequencyHz  := 60.0;
stMeas.fThdVoltsL1   := fThdVoltsPct;
stMeas.fThdVoltsL2   := fThdVoltsPct;
stMeas.fThdAmpsL1    := fThdAmpsPct;
stMeas.fThdAmpsL2    := fThdAmpsPct;

Read := bOnline;
END_METHOD

METHOD ReadHarmonics : BOOL
VAR_IN_OUT
    stHarm : ST_Harmonics;
END_VAR
VAR
    n : INT;
END_VAR
// A plausible switch-mode supply spectrum: odd orders falling off with the order, even orders near zero.
FOR n := 2 TO GVL_Param.HARMONIC_MAX_ORDER DO
    IF (n MOD 2) = 1 THEN
        stHarm.aAmpsL1[n]  := fThdAmpsPct * 2.2 / INT_TO_LREAL(n);
        stHarm.aVoltsL1[n] := fThdVoltsPct * 2.2 / INT_TO_LREAL(n);
    ELSE
        stHarm.aAmpsL1[n]  := 0.2;
        stHarm.aVoltsL1[n] := 0.1;
    END_IF
    stHarm.aAmpsL2[n]  := stHarm.aAmpsL1[n];
    stHarm.aVoltsL2[n] := stHarm.aVoltsL1[n];
END_FOR
stHarm.bValid := bOnline;

ReadHarmonics := bOnline;
END_METHOD

END_FUNCTION_BLOCK

// ---- POUs/Power/FB_SatelliteController.TcPOU
FUNCTION_BLOCK FB_SatelliteController IMPLEMENTS I_FeedLoad, I_JsonSource
VAR_INPUT
    stCfg : ST_BoxConfig;  // this box's row of GVL_Config.aBoxes
END_VAR
VAR_OUTPUT
    bValid      : BOOL;   // the values below can be used
    bMeasured   : BOOL;   // TRUE: from the supply. FALSE: estimated from the feed
    fDcAmps     : LREAL;  // A DC, filtered
    fDcVolts    : LREAL;  // V DC
    fAcPowerW   : LREAL;  // W on the AC side, at the box
    fCableLossW : LREAL;  // W lost in the box's own AC cable, on top of fAcPowerW
END_VAR
VAR
    fbSupply  : FB_EcPowerSupply;
    fEff      : LREAL := 0.95;
    fCycleS   : LREAL;
    fRawLossW : LREAL;  // cable loss from this cycle's unfiltered current
END_VAR

fEff    := LIMIT(0.5, stCfg.fPsuEfficiency, 1.0);
fCycleS := F_CycleTimeS();

IF stCfg.bHasEcPowerSupply THEN
    bMeasured := TRUE;
    fbSupply(bSimulate := GVL_Config.bSimulateSupplies);

    IF fbSupply.bOnline THEN
        fDcVolts  := fbSupply.fOutputVolts;
        // The loss goes with the square of the current, so it is taken from the raw current every cycle and
        // filtered afterwards. Filtering the current first would read low whenever the load moves.
        fRawLossW := F_CableLossW(fPowerW := fDcVolts * fbSupply.fOutputAmps / fEff,
                                  fLengthFt := stCfg.fWireLengthFt, nAwg := stCfg.nWireAwg);
        IF bValid THEN
            fDcAmps     := F_LowPass(fState := fDcAmps,     fInput := fbSupply.fOutputAmps, fTimeS := GVL_Config.fFilterTimeS, fCycleS := fCycleS);
            fCableLossW := F_LowPass(fState := fCableLossW, fInput := fRawLossW,            fTimeS := GVL_Config.fFilterTimeS, fCycleS := fCycleS);
        ELSE
            fDcAmps     := fbSupply.fOutputAmps;  // first valid sample: no filter run-in
            fCableLossW := fRawLossW;
        END_IF
        fAcPowerW := fDcVolts * fDcAmps / fEff;
        bValid    := TRUE;
    ELSE
        // Off the bus: counted as 0 W and reported as not valid.
        fDcAmps     := 0.0;
        fDcVolts    := 0.0;
        fAcPowerW   := 0.0;
        fCableLossW := 0.0;
        bValid      := FALSE;
    END_IF
ELSE
    // No supply: SetShare() writes the outputs when the feed has done its split.
    bMeasured := FALSE;
END_IF

METHOD GetDemand : ST_LoadDemand
VAR
    stDemand : ST_LoadDemand;
END_VAR
// What the feed sees at the branch point: the box's draw plus the loss in the box's cable.
stDemand.fCableFactor := F_CableFactor(fLengthFt := stCfg.fWireLengthFt, nAwg := stCfg.nWireAwg);
IF stCfg.bHasEcPowerSupply THEN
    stDemand.eKind       := E_LoadKind.Measured;
    stDemand.fAcPowerW   := fAcPowerW + fCableLossW;
    stDemand.fCableLossW := fCableLossW;
    stDemand.fWeight     := 0.0;
    stDemand.bValid      := bValid;
ELSE
    stDemand.eKind       := E_LoadKind.Estimated;
    stDemand.fAcPowerW   := 0.0;
    stDemand.fCableLossW := fCableLossW;  // from the share, once SetShare() has run this cycle
    stDemand.fWeight     := UDINT_TO_LREAL(stCfg.nPixelCount);
    stDemand.bValid      := TRUE;
END_IF
GetDemand := stDemand;
END_METHOD

METHOD SetShare
VAR_INPUT
    fShareW     : LREAL;  // W on the AC side
    bShareValid : BOOL;   // FALSE: the feed has no valid measurement
END_VAR
IF NOT stCfg.bHasEcPowerSupply THEN
    // The share includes the loss in the box's own cable. What arrives at the box is less.
    fAcPowerW   := F_PowerAfterCable(fShareW := fShareW, fLengthFt := stCfg.fWireLengthFt, nAwg := stCfg.nWireAwg);
    fCableLossW := MAX(0.0, fShareW) - fAcPowerW;
    fDcVolts    := stCfg.fNominalDcVolts;
    IF stCfg.fNominalDcVolts > 1.0 THEN
        fDcAmps := fAcPowerW * fEff / stCfg.fNominalDcVolts;
    ELSE
        fDcAmps := 0.0;
    END_IF
    bValid := bShareValid;
END_IF
END_METHOD

METHOD WriteJson
VAR_INPUT
    eSection : E_JsonSection;
END_VAR
VAR_IN_OUT
    fbJson : FB_JsonSaxWriter;
END_VAR
VAR
    sFeed : STRING(20);
END_VAR
IF eSection <> E_JsonSection.Box THEN
    RETURN;
END_IF

sFeed := F_FeedIdString(nFeedId := stCfg.nFeedId);

fbJson.AddKey('id');
fbJson.AddString(stCfg.sId);
fbJson.AddKey('name');
fbJson.AddString(stCfg.sControllerName);
fbJson.AddKey('feed');
fbJson.AddString(sFeed);
F_JsonInt(sKey := 'pixels', nValue := UDINT_TO_DINT(MIN(stCfg.nPixelCount, 2147483647)), fbJson := fbJson);
F_JsonNum(sKey := 'maxDcAmps', fValue := stCfg.fMaxDcCurrent, bValid := TRUE, nDecimals := 1, fbJson := fbJson);
fbJson.AddKey('src');
IF stCfg.bHasEcPowerSupply THEN
    fbJson.AddString('psu');
ELSE
    fbJson.AddString('est');
END_IF
fbJson.AddKey('ok');
fbJson.AddBool(bValid);
F_JsonNum(sKey := 'dcAmps', fValue := fDcAmps, bValid := bValid, nDecimals := 2, fbJson := fbJson);
F_JsonNum(sKey := 'dcVolts', fValue := fDcVolts, bValid := bValid AND stCfg.bHasEcPowerSupply, nDecimals := 1, fbJson := fbJson);
F_JsonNum(sKey := 'acW', fValue := fAcPowerW, bValid := bValid, nDecimals := 1, fbJson := fbJson);
F_JsonNum(sKey := 'cableLossW', fValue := fCableLossW, bValid := bValid, nDecimals := 1, fbJson := fbJson);

fbJson.AddKey('psu');
IF stCfg.bHasEcPowerSupply THEN
    fbJson.StartObject();
    fbJson.AddKey('dcOk');
    fbJson.AddBool(fbSupply.bDcOk);
    fbJson.AddKey('warn');
    fbJson.AddBool(fbSupply.bWarning);
    fbJson.AddKey('err');
    fbJson.AddBool(fbSupply.bError);
    F_JsonNumSigned(sKey := 'tempC', fValue := fbSupply.fTempC, bValid := fbSupply.bTempValid, nDecimals := 0, fbJson := fbJson);
    F_JsonNum(sKey := 'inVolts', fValue := fbSupply.fInputVolts, bValid := fbSupply.bInputVoltsValid, nDecimals := 0, fbJson := fbJson);
    fbJson.EndObject();
ELSE
    fbJson.AddNull();
END_IF
END_METHOD

END_FUNCTION_BLOCK

// ---- POUs/Power/FB_EcPowerSupply.TcPOU
FUNCTION_BLOCK FB_EcPowerSupply
VAR_INPUT
    bSimulate : BOOL;  // TRUE: use the fSim values below instead of the process image
END_VAR
VAR_OUTPUT
    bOnline          : BOOL;   // on the bus, in OP, data valid
    bDcOk            : BOOL;   // output voltage above the supply's DC OK threshold (22 V by default)
    bWarning         : BOOL;
    bError           : BOOL;
    fOutputVolts     : LREAL;  // V DC
    fOutputAmps      : LREAL;  // A DC
    bTempValid       : BOOL;
    fTempC           : LREAL;  // from info data 1
    bInputVoltsValid : BOOL;
    fInputVolts      : LREAL;  // V AC RMS, from info data 2
END_VAR
VAR
    // Process image. Linked in step 5.
    bInWarning       AT %I* : BOOL;  // 6000:01 Warning
    bInError         AT %I* : BOOL;  // 6000:02 Error
    bInDcOk          AT %I* : BOOL;  // 6000:04 DC OK
    fInOutputVoltage AT %I* : REAL;  // 6000:11 Output voltage, V
    fInOutputCurrent AT %I* : REAL;  // 6000:12 Output current, A
    nInInfoData1     AT %I* : UINT;  // 6000:15 Info data 1. Set 8001:19 = 14 (actual temperature)
    nInInfoData2     AT %I* : UINT;  // 6000:16 Info data 2. Set 8001:21 = 10 (actual RMS input voltage)
    bInWcState       AT %I* : BOOL;  // WcState. FALSE = data valid
    nInState         AT %I* : UINT;  // InfoData > State. 8 = OP

    // Simulation values. Change them online.
    fSimVolts      : LREAL := 24.0;
    fSimAmps       : LREAL := 5.0;
    fSimTempC      : LREAL := 35.0;
    fSimInputVolts : LREAL := 240.0;

    bFinite : BOOL;
    fVolts  : LREAL;
    fAmps   : LREAL;
END_VAR

IF bSimulate THEN
    bOnline          := TRUE;
    bDcOk            := TRUE;
    bWarning         := FALSE;
    bError           := FALSE;
    fOutputVolts     := fSimVolts;
    fOutputAmps      := fSimAmps;
    fTempC           := fSimTempC;
    fInputVolts      := fSimInputVolts;
    bTempValid       := TRUE;
    bInputVoltsValid := TRUE;
ELSE
    bFinite := TRUE;
    fVolts  := F_CleanReal(fIn := fInOutputVoltage, bAllFinite := bFinite);
    fAmps   := F_CleanReal(fIn := fInOutputCurrent, bAllFinite := bFinite);

    bOnline  := (nInState = 8) AND (NOT bInWcState) AND bFinite;
    // A supply that drops off the bus leaves its last values in the process image, so the bits only count while it is online.
    bDcOk    := bOnline AND bInDcOk;
    bWarning := bOnline AND bInWarning;
    bError   := bOnline AND bInError;

    IF bOnline THEN
        fOutputVolts := MAX(0.0, fVolts);
        fOutputAmps  := MAX(0.0, fAmps);
        fTempC       := INT_TO_LREAL(UINT_TO_INT(nInInfoData1)) * GVL_Config.fPsuInfo1Scale;  // read as signed: a box can be below 0 degrees C
        fInputVolts  := UINT_TO_LREAL(nInInfoData2) * GVL_Config.fPsuInfo2Scale;
    ELSE
        fOutputVolts := 0.0;
        fOutputAmps  := 0.0;
        fTempC       := 0.0;
        fInputVolts  := 0.0;
    END_IF
    bTempValid       := bOnline AND (GVL_Config.fPsuInfo1Scale > 0.0);
    bInputVoltsValid := bOnline AND (GVL_Config.fPsuInfo2Scale > 0.0);
END_IF

END_FUNCTION_BLOCK

// ---- POUs/Util/F_CleanReal.TcPOU
FUNCTION F_CleanReal : LREAL
VAR_INPUT
    fIn : REAL;
END_VAR
VAR_IN_OUT
    bAllFinite : BOOL;  // set FALSE when fIn is NaN or infinite; never set TRUE here
END_VAR
VAR
    fTmp : REAL;
END_VAR

fTmp := fIn;
IF IsFinite(F_REAL(fTmp)) THEN
    F_CleanReal := fTmp;
ELSE
    F_CleanReal := 0.0;
    bAllFinite := FALSE;
END_IF

END_FUNCTION

// ---- POUs/Util/F_CableLossW.TcPOU
FUNCTION F_CableLossW : LREAL
VAR_INPUT
    fPowerW   : LREAL;  // W at the load's terminals
    fLengthFt : LREAL;  // one-way length of its cable
    nAwg      : INT;
END_VAR
VAR
    fP : LREAL;
END_VAR

fP := MAX(0.0, fPowerW);
F_CableLossW := F_CableFactor(fLengthFt := fLengthFt, nAwg := nAwg) * fP * fP;

END_FUNCTION

// ---- POUs/Util/F_CableFactor.TcPOU
FUNCTION F_CableFactor : LREAL
VAR_INPUT
    fLengthFt : LREAL;  // one-way length of the cable
    nAwg      : INT;
END_VAR
VAR
    fVoltsEff : LREAL;  // V * PF
END_VAR

fVoltsEff := GVL_Config.fNominalAcVolts * LIMIT(0.5, GVL_Config.fNominalPowerFactor, 1.0);
IF fVoltsEff > 1.0 THEN
    F_CableFactor := 2.0 * F_WireOhms(fLengthFt := fLengthFt, nAwg := nAwg) / (fVoltsEff * fVoltsEff);
ELSE
    F_CableFactor := 0.0;
END_IF

END_FUNCTION

// ---- POUs/Util/F_PowerAfterCable.TcPOU
FUNCTION F_PowerAfterCable : LREAL
VAR_INPUT
    fShareW   : LREAL;  // W at the branch point
    fLengthFt : LREAL;  // one-way length of the cable
    nAwg      : INT;
END_VAR
VAR
    fA     : LREAL;
    fShare : LREAL;
END_VAR

fShare := MAX(0.0, fShareW);
fA     := F_CableFactor(fLengthFt := fLengthFt, nAwg := nAwg);
F_PowerAfterCable := 2.0 * fShare / (1.0 + SQRT(1.0 + 4.0 * fA * fShare));

END_FUNCTION

// ---- POUs/Util/F_FeedIdString.TcPOU
FUNCTION F_FeedIdString : STRING(20)
VAR_INPUT
    nFeedId : INT;
END_VAR

IF (nFeedId >= 1) AND (nFeedId <= GVL_Param.FEED_COUNT) THEN
    F_FeedIdString := GVL_Config.aFeeds[nFeedId].sId;
ELSE
    F_FeedIdString := '';
END_IF

END_FUNCTION

// ---- POUs/Util/F_JsonInt.TcPOU
FUNCTION F_JsonInt : BOOL
VAR_INPUT
    sKey   : STRING(31);
    nValue : DINT;
END_VAR
VAR_IN_OUT
    fbJson : FB_JsonSaxWriter;
END_VAR

fbJson.AddKey(sKey);
fbJson.AddDint(nValue);
F_JsonInt := TRUE;

END_FUNCTION

// ---- POUs/Power/FB_GenericLoad.TcPOU
FUNCTION_BLOCK FB_GenericLoad IMPLEMENTS I_FeedLoad, I_JsonSource
VAR_INPUT
    stCfg : ST_GenericLoadConfig;  // this load's row of GVL_Config.aLoads
END_VAR
VAR_OUTPUT
    fAcPowerW   : LREAL;  // W at the load
    fCableLossW : LREAL;  // W lost in the load's cable, on top of fAcPowerW
END_VAR

IF stCfg.bEnabled THEN
    fAcPowerW := MAX(0.0, stCfg.fRatedPowerW);
ELSE
    fAcPowerW := 0.0;
END_IF
fCableLossW := F_CableLossW(fPowerW := fAcPowerW, fLengthFt := stCfg.fWireLengthFt, nAwg := stCfg.nWireAwg);

METHOD GetDemand : ST_LoadDemand
VAR
    stDemand : ST_LoadDemand;
END_VAR
stDemand.eKind        := E_LoadKind.Rated;
stDemand.fAcPowerW    := fAcPowerW + fCableLossW;
stDemand.fCableLossW  := fCableLossW;
stDemand.fWeight      := 0.0;
stDemand.fCableFactor := F_CableFactor(fLengthFt := stCfg.fWireLengthFt, nAwg := stCfg.nWireAwg);
stDemand.bValid       := TRUE;
GetDemand := stDemand;
END_METHOD

METHOD SetShare
VAR_INPUT
    fShareW     : LREAL;
    bShareValid : BOOL;
END_VAR
// A rated load takes no share. The method exists because I_FeedLoad requires it.
;
END_METHOD

METHOD WriteJson
VAR_INPUT
    eSection : E_JsonSection;
END_VAR
VAR_IN_OUT
    fbJson : FB_JsonSaxWriter;
END_VAR
VAR
    sFeed : STRING(20);
END_VAR
IF eSection <> E_JsonSection.Load THEN
    RETURN;
END_IF

sFeed := F_FeedIdString(nFeedId := stCfg.nFeedId);

fbJson.AddKey('id');
fbJson.AddString(stCfg.sId);
fbJson.AddKey('name');
fbJson.AddString(stCfg.sName);
fbJson.AddKey('feed');
fbJson.AddString(sFeed);
F_JsonNum(sKey := 'ratedW', fValue := stCfg.fRatedPowerW, bValid := TRUE, nDecimals := 0, fbJson := fbJson);
fbJson.AddKey('on');
fbJson.AddBool(stCfg.bEnabled);
F_JsonNum(sKey := 'cableLossW', fValue := fCableLossW, bValid := TRUE, nDecimals := 1, fbJson := fbJson);
END_METHOD

END_FUNCTION_BLOCK

// ---- POUs/System/FB_ShowClock.TcPOU
FUNCTION_BLOCK FB_ShowClock
VAR_OUTPUT
    bValid    : BOOL;        // the clock looks set (year 2025 or later)
    sUtcIso   : STRING(30);  // 2026-12-04T23:15:02.000Z
    nLocalDay : UDINT;       // days since 1601-01-01 in local time
    stUtc     : TIMESTRUCT;
END_VAR
VAR
    nUtc     : T_FILETIME64;   // 100 ns ticks since 1601-01-01, UTC
    nLastUtc : T_FILETIME64;
    nLocal   : T_FILETIME64;
    fbTz     : FB_FileTime64ToTzSpecificLocalTime;
END_VAR

nUtc  := F_GetSystemTime();
stUtc := FILETIME64_TO_SYSTEMTIME(nUtc);

sUtcIso := F_PadNum(nValue := WORD_TO_UDINT(stUtc.wYear), nDigits := 4);
sUtcIso := CONCAT(sUtcIso, '-');
sUtcIso := CONCAT(sUtcIso, F_PadNum(nValue := WORD_TO_UDINT(stUtc.wMonth), nDigits := 2));
sUtcIso := CONCAT(sUtcIso, '-');
sUtcIso := CONCAT(sUtcIso, F_PadNum(nValue := WORD_TO_UDINT(stUtc.wDay), nDigits := 2));
sUtcIso := CONCAT(sUtcIso, 'T');
sUtcIso := CONCAT(sUtcIso, F_PadNum(nValue := WORD_TO_UDINT(stUtc.wHour), nDigits := 2));
sUtcIso := CONCAT(sUtcIso, ':');
sUtcIso := CONCAT(sUtcIso, F_PadNum(nValue := WORD_TO_UDINT(stUtc.wMinute), nDigits := 2));
sUtcIso := CONCAT(sUtcIso, ':');
sUtcIso := CONCAT(sUtcIso, F_PadNum(nValue := WORD_TO_UDINT(stUtc.wSecond), nDigits := 2));
sUtcIso := CONCAT(sUtcIso, '.');
sUtcIso := CONCAT(sUtcIso, F_PadNum(nValue := WORD_TO_UDINT(stUtc.wMilliseconds), nDigits := 3));
sUtcIso := CONCAT(sUtcIso, 'Z');

// The time-zone block expects a clock that runs on steadily. After a step (first cycle, NTP correction) it starts afresh.
IF (nUtc < nLastUtc) OR ((nUtc - nLastUtc) > ULINT#50000000) THEN  // backwards, or more than 5 s forwards
    fbTz.A_Reset();
END_IF
nLastUtc := nUtc;

fbTz(in := nUtc, tzInfo := GVL_Config.stTimeZone);
nLocal := fbTz.out;
nLocalDay := ULINT_TO_UDINT(nLocal / ULINT#864000000000);  // 100 ns ticks per day

bValid := stUtc.wYear >= 2025;

END_FUNCTION_BLOCK

// ---- POUs/Util/F_PadNum.TcPOU
FUNCTION F_PadNum : STRING(10)
VAR_INPUT
    nValue  : UDINT;
    nDigits : INT;  // 1..10
END_VAR
VAR
    sText : STRING(10);
END_VAR

sText := UDINT_TO_STRING(nValue);
WHILE (LEN(sText) < nDigits) AND (LEN(sText) < 10) DO
    sText := CONCAT('0', sText);
END_WHILE
F_PadNum := sText;

END_FUNCTION

// ---- POUs/System/FB_Telemetry.TcPOU
FUNCTION_BLOCK FB_Telemetry
VAR_INPUT
    bEnable        : BOOL := TRUE;
    stCfg          : ST_MqttConfig;
    sPassword      : STRING(63);  // empty = stay offline
    sTimestamp     : STRING(30);  // UTC, ISO 8601
    bSimulated     : BOOL;        // TRUE while any value comes from a simulation
    fTotalPowerW   : LREAL;       // sum of the feeds, W
    fTotalAmps     : LREAL;       // sum of the feeds, A
    fEnergyTodayWh : LREAL;       // sum of the feeds, Wh
END_VAR
VAR_OUTPUT
    bConnected        : BOOL;
    hrLastError       : HRESULT;  // last error reported by the MQTT client
    nPublishCount     : UDINT;
    nDropCount        : UDINT;    // payload did not fit the buffer, or the client refused it
    nLastPayloadBytes : UDINT;
END_VAR
VAR
    fbMqtt : FB_IotMqttClient;
    fbJson : FB_JsonSaxWriter;
    sJson  : STRING(32000);       // payload buffer. Room for 64 boxes; the website drops anything above 64 KB

    // Sources handed in by MAIN this cycle
    aFeedSrc  : ARRAY[1..GVL_Param.FEED_COUNT] OF I_JsonSource;
    aBoxSrc   : ARRAY[1..GVL_Param.BOX_COUNT] OF I_JsonSource;
    aLoadSrc  : ARRAY[1..GVL_Param.LOAD_COUNT] OF I_JsonSource;
    ipDiagSrc : I_JsonSource;
    nFeedSrc  : INT;
    nBoxSrc   : INT;
    nLoadSrc  : INT;

    sTopicOnline : STRING(255);
    sTopicDash   : STRING(255);
    sTopicDiag   : STRING(255);
    sTopicHarm   : STRING(255);
    sOnline      : STRING(1) := '1';
    sOffline     : STRING(1) := '0';

    tonDash  : TON;
    tonDiag  : TON;
    tonHarm  : TON;
    bDashDue : BOOL;
    bDiagDue : BOOL;
    bHarmDue : BOOL;

    bRun          : BOOL;
    sPasswordSeen : STRING(63);
    bWasConnected : BOOL;
    bSendOnline   : BOOL;
    i             : INT;
END_VAR

// ---- topics ---------------------------------------------------------------
sTopicOnline := CONCAT(stCfg.sTopicRoot, '/online');
sTopicDash   := CONCAT(stCfg.sTopicRoot, '/dashboard');
sTopicDiag   := CONCAT(stCfg.sTopicRoot, '/diag');
sTopicHarm   := CONCAT(stCfg.sTopicRoot, '/harmonics');

// ---- connection. The client reads these settings when it connects -----------
fbMqtt.sHostName     := stCfg.sHost;
fbMqtt.nHostPort     := stCfg.nPort;
fbMqtt.sClientId     := stCfg.sClientId;
fbMqtt.sUserName     := stCfg.sUser;
fbMqtt.sUserPassword := sPassword;
fbMqtt.sTopicPrefix  := '';
fbMqtt.nKeepAlive    := stCfg.nKeepAliveS;

// Last will: the broker publishes "0" for us if the PLC drops off the network.
fbMqtt.stWill.sTopic       := sTopicOnline;
fbMqtt.stWill.pPayload     := ADR(sOffline);
fbMqtt.stWill.nPayloadSize := 1;
fbMqtt.stWill.eQoS         := TcIotMqttQos.AtLeastOnceDelivery;
fbMqtt.stWill.bRetain      := TRUE;

// A changed password drops the connection for one cycle, so the next attempt uses the new one.
bRun := bEnable AND stCfg.bEnable AND (LEN(sPassword) > 0) AND (sPassword = sPasswordSeen);
sPasswordSeen := sPassword;
fbMqtt.Execute(bRun);
bConnected := fbMqtt.bConnected;
IF fbMqtt.bError THEN
    hrLastError := fbMqtt.hrErrorCode;
END_IF

// ---- "online" once per connection --------------------------------------------
IF bConnected AND NOT bWasConnected THEN
    bSendOnline := TRUE;
    bDashDue    := TRUE;  // first frame right away
    hrLastError := 0;     // connected: the errors of the attempts before are history
END_IF
bWasConnected := bConnected;

IF bConnected AND bSendOnline THEN
    IF fbMqtt.Publish(sTopic := sTopicOnline, pPayload := ADR(sOnline), nPayloadSize := 1,
                      eQoS := TcIotMqttQos.AtLeastOnceDelivery, bRetain := TRUE, bQueue := FALSE) THEN
        bSendOnline := FALSE;
    END_IF
END_IF

// ---- timers ---------------------------------------------------------------------
tonDash(IN := bConnected AND NOT tonDash.Q, PT := stCfg.tDashboard);
IF tonDash.Q THEN
    bDashDue := TRUE;
END_IF
tonDiag(IN := bConnected AND NOT tonDiag.Q, PT := stCfg.tDiag);
IF tonDiag.Q THEN
    bDiagDue := TRUE;
END_IF
tonHarm(IN := bConnected AND NOT tonHarm.Q, PT := stCfg.tHarmonics);
IF tonHarm.Q THEN
    bHarmDue := TRUE;
END_IF
IF NOT bConnected THEN
    bDashDue := FALSE;
    bDiagDue := FALSE;
    bHarmDue := FALSE;
END_IF

// ---- one payload per cycle at most ------------------------------------------------
IF bDashDue THEN
    bDashDue := FALSE;

    fbJson.ResetDocument();
    fbJson.SetMaxDecimalPlaces(3);
    fbJson.StartObject();
    F_JsonInt(sKey := 'v', nValue := 2, fbJson := fbJson);
    fbJson.AddKey('ts');
    fbJson.AddString(sTimestamp);
    fbJson.AddKey('sim');
    fbJson.AddBool(bSimulated);
    // The three totals are required numbers in the website's original schema.
    F_JsonNum(sKey := 'powerW',        fValue := fTotalPowerW,   bValid := TRUE, nDecimals := 1, fbJson := fbJson);
    F_JsonNum(sKey := 'energyTodayWh', fValue := fEnergyTodayWh, bValid := TRUE, nDecimals := 0, fbJson := fbJson);
    F_JsonNum(sKey := 'totalAmps',     fValue := fTotalAmps,     bValid := TRUE, nDecimals := 2, fbJson := fbJson);

    fbJson.AddKey('circuits');
    fbJson.StartArray();
    FOR i := 1 TO nFeedSrc DO
        fbJson.StartObject();
        aFeedSrc[i].WriteJson(eSection := E_JsonSection.Circuit, fbJson := fbJson);
        fbJson.EndObject();
    END_FOR
    fbJson.EndArray();

    fbJson.AddKey('feeds');
    fbJson.StartArray();
    FOR i := 1 TO nFeedSrc DO
        fbJson.StartObject();
        aFeedSrc[i].WriteJson(eSection := E_JsonSection.Feed, fbJson := fbJson);
        fbJson.EndObject();
    END_FOR
    fbJson.EndArray();

    fbJson.AddKey('boxes');
    fbJson.StartArray();
    FOR i := 1 TO nBoxSrc DO
        fbJson.StartObject();
        aBoxSrc[i].WriteJson(eSection := E_JsonSection.Box, fbJson := fbJson);
        fbJson.EndObject();
    END_FOR
    fbJson.EndArray();

    fbJson.AddKey('loads');
    fbJson.StartArray();
    FOR i := 1 TO nLoadSrc DO
        fbJson.StartObject();
        aLoadSrc[i].WriteJson(eSection := E_JsonSection.Load, fbJson := fbJson);
        fbJson.EndObject();
    END_FOR
    fbJson.EndArray();

    fbJson.EndObject();
    Send(sTopic := sTopicDash);

ELSIF bDiagDue THEN
    bDiagDue := FALSE;

    IF ipDiagSrc <> 0 THEN
        fbJson.ResetDocument();
        fbJson.SetMaxDecimalPlaces(3);
        fbJson.StartObject();
        ipDiagSrc.WriteJson(eSection := E_JsonSection.Diag, fbJson := fbJson);
        fbJson.EndObject();
        Send(sTopic := sTopicDiag);
    END_IF

ELSIF bHarmDue THEN
    bHarmDue := FALSE;

    IF nFeedSrc > 0 THEN
        fbJson.ResetDocument();
        fbJson.SetMaxDecimalPlaces(3);
        fbJson.StartObject();
        fbJson.AddKey('ts');
        fbJson.AddString(sTimestamp);
        fbJson.AddKey('feeds');
        fbJson.StartArray();
        FOR i := 1 TO nFeedSrc DO
            fbJson.StartObject();
            aFeedSrc[i].WriteJson(eSection := E_JsonSection.Harmonics, fbJson := fbJson);
            fbJson.EndObject();
        END_FOR
        fbJson.EndArray();
        fbJson.EndObject();
        Send(sTopic := sTopicHarm);
    END_IF
END_IF

// ---- MAIN hands the sources in again next cycle -------------------------------------
nFeedSrc  := 0;
nBoxSrc   := 0;
nLoadSrc  := 0;
ipDiagSrc := 0;

// Call every cycle, before the block itself, once per object that should appear in the payloads.
METHOD AddSource : BOOL
VAR_INPUT
    eSection : E_JsonSection;  // Feed, Box, Load or Diag
    ipSource : I_JsonSource;
END_VAR
AddSource := FALSE;
IF ipSource = 0 THEN
    RETURN;
END_IF

CASE eSection OF
    E_JsonSection.Feed:
        IF nFeedSrc < GVL_Param.FEED_COUNT THEN
            nFeedSrc := nFeedSrc + 1;
            aFeedSrc[nFeedSrc] := ipSource;
            AddSource := TRUE;
        END_IF
    E_JsonSection.Box:
        IF nBoxSrc < GVL_Param.BOX_COUNT THEN
            nBoxSrc := nBoxSrc + 1;
            aBoxSrc[nBoxSrc] := ipSource;
            AddSource := TRUE;
        END_IF
    E_JsonSection.Load:
        IF nLoadSrc < GVL_Param.LOAD_COUNT THEN
            nLoadSrc := nLoadSrc + 1;
            aLoadSrc[nLoadSrc] := ipSource;
            AddSource := TRUE;
        END_IF
    E_JsonSection.Diag:
        ipDiagSrc := ipSource;
        AddSource := TRUE;
END_CASE
END_METHOD

// Publishes the document the JSON writer holds. QoS 1, retained, no trailing zero byte.
METHOD PRIVATE Send : BOOL
VAR_INPUT
    sTopic : STRING(255);
END_VAR
VAR
    nLen  : UDINT;
    bSent : BOOL;
END_VAR
bSent := FALSE;
nLen := fbJson.CopyDocument(sJson, SIZEOF(sJson));  // length including the terminating zero; 0 = did not fit
IF nLen > 1 THEN
    nLastPayloadBytes := nLen - 1;
    bSent := fbMqtt.Publish(sTopic := sTopic, pPayload := ADR(sJson), nPayloadSize := nLen - 1,
                            eQoS := TcIotMqttQos.AtLeastOnceDelivery, bRetain := TRUE, bQueue := FALSE);
END_IF

IF bSent THEN
    nPublishCount := nPublishCount + 1;
ELSE
    nDropCount := nDropCount + 1;
END_IF
Send := bSent;
END_METHOD

END_FUNCTION_BLOCK

// ---- POUs/System/FB_IpcDiagnostics.TcPOU
FUNCTION_BLOCK FB_IpcDiagnostics IMPLEMENTS I_JsonSource
VAR_INPUT
    bEnable : BOOL := TRUE;  // FALSE: leave the Device Manager alone
	sHostThermalPath : STRING(255) := '/sys/class/hwmon/hwmon2/temp2_input';  // Zynq FPD: the A53 cores. hwmon1 = rv3032 RTC (board), hwmon2 temp1 = LPD
END_VAR
VAR_OUTPUT
    // PLC task
    nCycleUs     : UDINT;    // configured cycle time
    nLastExecUs  : UDINT;    // execution time of the last cycle
    nExceedCount : UDINT;    // cycles that overran since the PLC started
    fUptimeS     : LREAL;    // PLC run time
    bRtCpuValid  : BOOL;
    fRtCpuPct    : LREAL;    // TwinCAT real-time share of the CPU

    // Controller, from the Device Manager
    bMdpReady    : BOOL;     // the Device Manager answered
    hrMdpError   : HRESULT;  // last error from registration or a read
    bCpuValid    : BOOL;
    fCpuPct      : LREAL;    // whole-controller CPU load
    bTempValid   : BOOL;
    fCpuTempC    : LREAL;
    bMemValid    : BOOL;
    fMemPct      : LREAL;    // RAM in use
    bDiskValid   : BOOL;
    fDiskPct     : LREAL;    // storage in use, largest volume

    // EtherCAT master
    bEcLinked    : BOOL;     // the three inputs below are linked
    bEcOk        : BOOL;
END_VAR
VAR
    // Optional links to the EtherCAT master (step 3)
    nEcDevState   AT %I* : UINT;  // Inputs > DevState. 0 = no fault
    nEcSlaveCount AT %I* : UINT;  // Inputs > SlaveCount: slaves found
    nEcCfgSlaves  AT %I* : UINT;  // InfoData > CfgSlaveCount: slaves configured

    nTaskIdx : DINT;

    // TwinCAT real-time share
    fbRtCpu  : TC_CpuUsage;
    tonRtCpu : TON;
    nRtStep  : INT;

    // Kernel temperature
    fbThermal  : FB_HostThermal;
    bMdpTemp   : BOOL;   // the Device Manager served CPU_Temp in the last round

    // Device Manager
    fbRegister : FB_IPCDiag_Register;
    fbRead     : FB_IPCDiag_ReadParameter;
    tonMdp     : TON;
    nMdpStep   : INT;
    nKey       : INT;
    aKeys      : ARRAY[1..KEY_COUNT] OF E_IPCDiag_ParameterKey := [
                     E_IPCDiag_ParameterKey.CPU_Usage,
                     E_IPCDiag_ParameterKey.CPU_Temp,
                     E_IPCDiag_ParameterKey.Memory_ProgramMemoryAllocated,
                     E_IPCDiag_ParameterKey.Memory_ProgramMemoryAvailable,
                     E_IPCDiag_ParameterKey.Disk_VolumeList_TotelSize,
                     E_IPCDiag_ParameterKey.Disk_VolumeList_FreeSpace];
    hr         : HRESULT;
    nValU16    : UINT;
    nValI16    : INT;
    nValU64    : ULINT;
    nMemTotal  : ULINT;
    bMemTotOk  : BOOL;
    aVolTotal  : ARRAY[1..MAX_VOLUMES] OF ULINT;
    nVolCount  : USINT;
    nFreeCount : USINT;
    nBest      : USINT;
    nBestSize  : ULINT;
    j          : USINT;
END_VAR
VAR CONSTANT
    KEY_COUNT   : INT := 6;
    MAX_VOLUMES : USINT := 8;
END_VAR

// ---- PLC task ---------------------------------------------------------------
nTaskIdx := GETCURTASKINDEXEX();
IF (nTaskIdx >= 1) AND (nTaskIdx <= 20) THEN
    nCycleUs    := _TaskInfo[nTaskIdx].CycleTime / 10;     // 100 ns to microseconds
    nLastExecUs := _TaskInfo[nTaskIdx].LastExecTime / 10;
    IF _TaskInfo[nTaskIdx].CycleTimeExceeded THEN
        nExceedCount := nExceedCount + 1;
    END_IF
END_IF
fUptimeS := fUptimeS + F_CycleTimeS();

// ---- TwinCAT real-time share, every 5 s -------------------------------------------
CASE nRtStep OF
    0:
        tonRtCpu(IN := TRUE, PT := T#5S);
        IF tonRtCpu.Q THEN
            tonRtCpu(IN := FALSE);
            fbRtCpu(NETID := '', START := FALSE);
            fbRtCpu(NETID := '', START := TRUE, TMOUT := T#2S);
            nRtStep := 1;
        END_IF
    1:
        fbRtCpu(START := FALSE);
        IF NOT fbRtCpu.BUSY THEN
            bRtCpuValid := NOT fbRtCpu.ERR;
            IF bRtCpuValid THEN
                fRtCpuPct := UDINT_TO_LREAL(fbRtCpu.USAGE);
            END_IF
            nRtStep := 0;
        END_IF
ELSE
    nRtStep := 0;
END_CASE

// ---- Kernel temperature, every 10 s. The Device Manager on RT Linux has no CPU_Temp (V3) ---
fbThermal(bEnable := bEnable AND (LEN(sHostThermalPath) > 0), sPath := sHostThermalPath);

// ---- Device Manager: register once, then read one parameter after the other ----------
CASE nMdpStep OF
    0:  // the Device Manager needs time after boot
        tonMdp(IN := bEnable, PT := T#30S);
        IF tonMdp.Q THEN
            tonMdp(IN := FALSE);
            fbRegister(bExecute := FALSE);
            fbRegister(bExecute := TRUE);
            nMdpStep := 1;
        END_IF

    1:  // wait for the registration
        fbRegister(bExecute := FALSE);
        IF NOT fbRegister.bBusy THEN
            IF fbRegister.bError THEN
                hrMdpError := fbRegister.hrErrorCode;
                bMdpReady  := FALSE;
                nMdpStep   := 0;  // try again in 30 s
            ELSE
                bMdpReady := TRUE;
                nKey      := 1;
                nMdpStep  := 2;
            END_IF
        END_IF

    2:  // start one read
        fbRead(bExecute := FALSE, fbRegister := fbRegister);
        fbRead(bExecute := TRUE, eParameterKey := aKeys[nKey], fbRegister := fbRegister);
        nMdpStep := 3;

    3:  // wait for it, then take the value
        fbRead(bExecute := FALSE, fbRegister := fbRegister);
        IF NOT fbRead.bBusy THEN
            IF fbRead.bError THEN
                hrMdpError := fbRead.hrErrorCode;
            END_IF

            CASE nKey OF
                1:  // CPU load, UINT, %
                    bCpuValid := FALSE;
                    IF NOT fbRead.bError THEN
                        hr := fbRead.GetParameter(pBuffer := ADR(nValU16), nBufferSize := SIZEOF(nValU16));
                        IF SUCCEEDED(hr) THEN
                            fCpuPct   := LIMIT(0.0, UINT_TO_LREAL(nValU16), 100.0);
                            bCpuValid := TRUE;
                        END_IF
                    END_IF

                2:  // CPU temperature, INT, degrees C
                    bMdpTemp := FALSE;
                    IF fbRead.bError AND (nKey <> 2) THEN   // key 2 (CPU_Temp) has the kernel as fallback; its absence is not a faultN
                        hr := fbRead.GetParameter(pBuffer := ADR(nValI16), nBufferSize := SIZEOF(nValI16));
                        IF SUCCEEDED(hr) THEN
                            fCpuTempC  := INT_TO_LREAL(nValI16);
                            bMdpTemp := TRUE;
                        END_IF
                    END_IF

                3:  // RAM allocated, ULINT, bytes
                    bMemTotOk := FALSE;
                    IF NOT fbRead.bError THEN
                        hr := fbRead.GetParameter(pBuffer := ADR(nValU64), nBufferSize := SIZEOF(nValU64));
                        IF SUCCEEDED(hr) THEN
                            nMemTotal := nValU64;
                            bMemTotOk := nValU64 > 0;
                        END_IF
                    END_IF

                4:  // RAM available, ULINT, bytes
                    bMemValid := FALSE;
                    IF bMemTotOk AND NOT fbRead.bError THEN
                        hr := fbRead.GetParameter(pBuffer := ADR(nValU64), nBufferSize := SIZEOF(nValU64));
                        IF SUCCEEDED(hr) THEN
                            IF nValU64 <= nMemTotal THEN
                                fMemPct   := (1.0 - ULINT_TO_LREAL(nValU64) / ULINT_TO_LREAL(nMemTotal)) * 100.0;
                                bMemValid := TRUE;
                            END_IF
                        END_IF
                    END_IF

                5:  // total size of every volume, list of ULINT, bytes
                    nVolCount := 0;
                    IF NOT fbRead.bError THEN
                        nVolCount := MIN(fbRead.nReadParameterValues, MAX_VOLUMES);
                        FOR j := 1 TO nVolCount DO
                            hr := fbRead.GetParameterByIdx(pBuffer := ADR(nValU64), nBufferSize := SIZEOF(nValU64), nParameterIdx := j);
                            IF SUCCEEDED(hr) THEN
                                aVolTotal[j] := nValU64;
                            ELSE
                                aVolTotal[j] := 0;
                            END_IF
                        END_FOR
                    END_IF

                6:  // free space of every volume. The largest volume is taken as the system storage.
                    bDiskValid := FALSE;
                    IF (nVolCount > 0) AND NOT fbRead.bError THEN
                        nFreeCount := MIN(fbRead.nReadParameterValues, MAX_VOLUMES);
                        nBest     := 0;
                        nBestSize := 0;
                        FOR j := 1 TO nVolCount DO
                            IF aVolTotal[j] > nBestSize THEN
                                nBestSize := aVolTotal[j];
                                nBest     := j;
                            END_IF
                        END_FOR
                        IF (nBest >= 1) AND (nBest <= nFreeCount) THEN
                            hr := fbRead.GetParameterByIdx(pBuffer := ADR(nValU64), nBufferSize := SIZEOF(nValU64), nParameterIdx := nBest);
                            IF SUCCEEDED(hr) THEN
                                IF nValU64 <= nBestSize THEN
                                    fDiskPct   := (1.0 - ULINT_TO_LREAL(nValU64) / ULINT_TO_LREAL(nBestSize)) * 100.0;
                                    bDiskValid := TRUE;
                                END_IF
                            END_IF
                        END_IF
                    END_IF
            END_CASE

            IF nKey >= KEY_COUNT THEN
                nKey     := 1;
                nMdpStep := 4;
            ELSE
                nKey     := nKey + 1;
                nMdpStep := 2;
            END_IF
        END_IF

    4:  // pause between rounds
        tonMdp(IN := TRUE, PT := T#5S);
        IF tonMdp.Q THEN
            tonMdp(IN := FALSE);
            IF bEnable THEN
                nMdpStep := 2;
            END_IF
        END_IF
ELSE
    nMdpStep := 0;
END_CASE

// ---- Temperature: the Device Manager's CPU_Temp when it serves one, else the kernel's thermal zone ----
IF (NOT bMdpTemp) AND fbThermal.bValid THEN
    fCpuTempC := fbThermal.fTempC;
END_IF
bTempValid := bMdpTemp OR fbThermal.bValid;

// ---- EtherCAT master -------------------------------------------------------------------
bEcLinked := nEcCfgSlaves > 0;
bEcOk     := bEcLinked AND (nEcDevState = 0) AND (nEcSlaveCount = nEcCfgSlaves);

METHOD WriteJson
VAR_INPUT
    eSection : E_JsonSection;
END_VAR
VAR_IN_OUT
    fbJson : FB_JsonSaxWriter;
END_VAR
VAR
    fRt : LREAL;
END_VAR
IF eSection <> E_JsonSection.Diag THEN
    RETURN;
END_IF

// The first six keys are the website's original diag schema. They are required numbers there, so unknown is sent as 0.
fRt := 0.0;
IF bRtCpuValid THEN
    fRt := LIMIT(0.0, fRtCpuPct, 100.0);
END_IF
fbJson.AddKey('plcState');
fbJson.AddString('Run');
F_JsonNum(sKey := 'cpuPct', fValue := fRt, bValid := TRUE, nDecimals := 0, fbJson := fbJson);
F_JsonInt(sKey := 'cycleUs',     nValue := UDINT_TO_DINT(MIN(nCycleUs, 2147483647)),     fbJson := fbJson);
F_JsonInt(sKey := 'lastExecUs',  nValue := UDINT_TO_DINT(MIN(nLastExecUs, 2147483647)),  fbJson := fbJson);
F_JsonInt(sKey := 'exceedCount', nValue := UDINT_TO_DINT(MIN(nExceedCount, 2147483647)), fbJson := fbJson);
F_JsonNum(sKey := 'uptimeSec', fValue := fUptimeS, bValid := TRUE, nDecimals := 0, fbJson := fbJson);

fbJson.AddKey('ipc');
fbJson.StartObject();
F_JsonNum(sKey := 'cpuPct', fValue := fCpuPct, bValid := bCpuValid, nDecimals := 0, fbJson := fbJson);
F_JsonNumSigned(sKey := 'cpuTempC', fValue := fCpuTempC, bValid := bTempValid, nDecimals := 0, fbJson := fbJson);
F_JsonNum(sKey := 'memPct', fValue := fMemPct, bValid := bMemValid, nDecimals := 1, fbJson := fbJson);
F_JsonNum(sKey := 'diskPct', fValue := fDiskPct, bValid := bDiskValid, nDecimals := 1, fbJson := fbJson);
fbJson.EndObject();

fbJson.AddKey('ecat');
IF bEcLinked THEN
    fbJson.StartObject();
    fbJson.AddKey('ok');
    fbJson.AddBool(bEcOk);
    F_JsonInt(sKey := 'slaves',    nValue := UINT_TO_DINT(nEcSlaveCount), fbJson := fbJson);
    F_JsonInt(sKey := 'slavesCfg', nValue := UINT_TO_DINT(nEcCfgSlaves),  fbJson := fbJson);
    fbJson.EndObject();
ELSE
    fbJson.AddNull();
END_IF
END_METHOD

END_FUNCTION_BLOCK
